(* IEC 61131-3 sources: SortJet_MasterSPS_Aufbau.fbsproj/09_Station/UnterStationsbausteine/Entwicklung/Motorstarter_FB_V01_00_00.fb.st^, 4 files *)

(* ---- A_Changelog.act.st ---- *)
(* METADATA
{
	"v3Meta": {
		"objectGuid": "e9ea620c-f297-40f4-a2c5-b8d2a96a7ee4"
	}
}
*)
{attribute 'excludefrombuild'}
ACTION A_Changelog
(* !!! VERSIONSÄNDERUNGEN WERDEN HIER DETAILLIERT DOKUMENTIERT !!!

- 2026-11-24 - V01_00_00: Tobias Brekerbohm
  - Erste Freigabe SortJet-Master
*)
END_ACTION

(* ---- Linkslauf.meth.st ---- *)
(* METADATA
{
	"v3Meta": {
		"objectGuid": "901ae501-1a81-4a6e-8340-32118915e16c"
	}
}
*)
METHOD Linkslauf : BOOL
VAR_INPUT
END_VAR

VAR
  tonlMaxWarteZeit : TON;

END_VAR
Linkslauf := FALSE;

tonlMaxWarteZeit( IN := TRUE, PT:= T#4000MS );
IF ( tonlMaxWarteZeit.Q ) THEN
  bpFehler := TRUE;
  wpFehlerNr := cMELDUNG_MOTORSTARTER_FEHLER_LINKSLAUF_OK;
  out_bLinkslauf := FALSE;
END_IF

out_bLinkslauf := bpSensorNotNockeLinkslauf;

IF NOT bpSensorNotNockeLinkslauf THEN
  Linkslauf := TRUE;
END_IF
END_METHOD

(* ---- Rechtslauf.meth.st ---- *)
(* METADATA
{
	"v3Meta": {
		"objectGuid": "9a97d710-cc7f-4070-b236-0ffc8d0344e1"
	}
}
*)
METHOD Rechtslauf : BOOL
VAR_INPUT
END_VAR

VAR
  tonlMaxWarteZeit : TON;

END_VAR
Rechtslauf := FALSE;

tonlMaxWarteZeit( IN := TRUE, PT:= T#4000MS );
IF ( tonlMaxWarteZeit.Q )THEN
  bpFehler := TRUE;
  wpFehlerNr := cMELDUNG_MOTORSTARTER_FEHLER_RECHTSLAUF_OK;
  out_bRechtslauf := FALSE;
END_IF

out_bRechtslauf := bpSensorNotNockeRechtslauf;

IF NOT bpSensorNotNockeRechtslauf THEN
  Rechtslauf := TRUE;
END_IF
END_METHOD

(* ---- Reset.meth.st ---- *)
(* METADATA
{
	"v3Meta": {
		"objectGuid": "5e136676-7d5d-430e-b251-8802f4b156e4"
	}
}
*)
METHOD Reset : BOOL
VAR_INPUT

END_VAR

VAR
  tonlReset : TON;

END_VAR

tonlReset( IN := TRUE , PT :=  T#1500MS );
out_Reset := NOT tonlReset.Q;

Reset := bpMotorstarterOK;
END_METHOD
